(* IEC 61131-3 sources: 2026_Projet_YGO_ExcavatriceDragage/CODE_BACKUP/CODE_20260822_IntroductionTestCI/J_SUPERVISION/_BRIDGES, 7 files *)

(* ---- FB_CfgPersistBridge_BucketCfg.st ---- *)
(* =======================================================================
   💾 FB_CfgPersistBridge_BucketCfg — Pont persistance pour ST_BucketCfg
   ───────────────────────────────────────────────────────────────
   🎯 Rôle : Restauration et synchronisation bidirectionnelle IHM / Persist
   💾 Persistance : Transfert GVL_PERSISTENT <-> GVL_IHM sur Initialized
   📄 Doc métier : DOC/AF/AF_Partie-03_Contrats_Composants_v2.1.md §3
   ======================================================================= *)
FUNCTION_BLOCK FB_CfgPersistBridge_BucketCfg
VAR_OUTPUT
    // === ETATS RESTAURATION ===
    JustRestored            : BOOL;               // <-- [STAT] Vrai sur le cycle de restauration initiale
END_VAR
VAR_IN_OUT
    // === BUS CONFIGURATION ET PERSISTANCE ===
    Hmi                     : ST_BucketCfg;       // <-> [BUS] Structure de configuration IHM
    Persist                 : ST_BucketCfg;       // <-> [BUS] Structure de configuration persistante
END_VAR

JustRestored := FALSE;
IF NOT Hmi.Initialized THEN
    Hmi := Persist;
    Hmi.Initialized := TRUE;
    JustRestored := TRUE;
ELSE
    Persist := Hmi;
END_IF;

(* ---- FB_CfgPersistBridge_CommunCfg.st ---- *)
(* =======================================================================
   💾 FB_CfgPersistBridge_CommunCfg — Pont persistance pour ST_CommunCfg
   ───────────────────────────────────────────────────────────────
   🎯 Rôle : Restauration et synchronisation bidirectionnelle IHM / Persist
   💾 Persistance : Transfert GVL_PERSISTENT <-> GVL_IHM sur Initialized
   📄 Doc métier : DOC/AF/AF_Partie-03_Contrats_Composants_v2.1.md §3
   ======================================================================= *)
FUNCTION_BLOCK FB_CfgPersistBridge_CommunCfg
VAR_OUTPUT
    // === ETATS RESTAURATION ===
    JustRestored            : BOOL;               // <-- [STAT] Vrai sur le cycle de restauration initiale
END_VAR
VAR_IN_OUT
    // === BUS CONFIGURATION ET PERSISTANCE ===
    Hmi                     : ST_CommunCfg;       // <-> [BUS] Structure de configuration IHM
    Persist                 : ST_CommunCfg;       // <-> [BUS] Structure de configuration persistante
END_VAR

JustRestored := FALSE;
IF NOT Hmi.Initialized THEN
    Hmi := Persist;
    Hmi.Initialized := TRUE;
    JustRestored := TRUE;
ELSE
    Persist := Hmi;
END_IF;

(* ---- FB_CfgPersistBridge_CycleCfg.st ---- *)
(* =======================================================================
   💾 FB_CfgPersistBridge_CycleCfg — Pont persistance pour ST_CycleCfg
   ───────────────────────────────────────────────────────────────
   🎯 Rôle : Restauration et synchronisation bidirectionnelle IHM / Persist
   💾 Persistance : Transfert GVL_PERSISTENT <-> GVL_IHM sur Initialized
   📄 Doc métier : DOC/AF/AF_Partie-03_Contrats_Composants_v2.1.md §3
   ======================================================================= *)
FUNCTION_BLOCK FB_CfgPersistBridge_CycleCfg
VAR_OUTPUT
    // === ETATS RESTAURATION ===
    JustRestored            : BOOL;               // <-- [STAT] Vrai sur le cycle de restauration initiale
END_VAR
VAR_IN_OUT
    // === BUS CONFIGURATION ET PERSISTANCE ===
    Hmi                     : ST_CycleCfg;        // <-> [BUS] Structure de configuration IHM
    Persist                 : ST_CycleCfg;        // <-> [BUS] Structure de configuration persistante
END_VAR

JustRestored := FALSE;
IF NOT Hmi.Initialized THEN
    Hmi := Persist;
    Hmi.Initialized := TRUE;
    JustRestored := TRUE;
ELSE
    Persist := Hmi;
END_IF;

(* ---- FB_CfgPersistBridge_DredgingAssistCfg.st ---- *)
(* =======================================================================
   💾 FB_CfgPersistBridge_DredgingAssistCfg — Pont persistance prélèvement
   ───────────────────────────────────────────────────────────────
   🎯 Rôle : Restauration et synchronisation bidirectionnelle IHM / Persist
   💾 Persistance : Transfert GVL_PERSISTENT <-> GVL_IHM sur Initialized
   📄 Doc métier : DOC/AF/AF_Partie-03_Contrats_Composants_v2.1.md §3
   ======================================================================= *)
FUNCTION_BLOCK FB_CfgPersistBridge_DredgingAssistCfg
VAR_OUTPUT
    // === ETATS RESTAURATION ===
    JustRestored            : BOOL;               // <-- [STAT] Vrai sur le cycle de restauration initiale
END_VAR
VAR_IN_OUT
    // === BUS CONFIGURATION ET PERSISTANCE ===
    Hmi                     : ST_DredgingAssistCfg; // <-> [BUS] Structure de configuration IHM
    Persist                 : ST_DredgingAssistCfg; // <-> [BUS] Structure de configuration persistante
END_VAR

JustRestored := FALSE;
IF NOT Hmi.Initialized THEN
    Hmi := Persist;
    Hmi.Initialized := TRUE;
    JustRestored := TRUE;
ELSE
    Persist := Hmi;
END_IF;

(* ---- FB_CfgPersistBridge_SyncCfg.st ---- *)
(* =======================================================================
   💾 FB_CfgPersistBridge_SyncCfg — Pont persistance pour ST_SyncCfg
   ───────────────────────────────────────────────────────────────
   🎯 Rôle : Restauration et synchronisation bidirectionnelle IHM / Persist
   💾 Persistance : Transfert GVL_PERSISTENT <-> GVL_IHM sur Initialized
   📄 Doc métier : DOC/AF/AF_Partie-03_Contrats_Composants_v2.1.md §3
   ======================================================================= *)
FUNCTION_BLOCK FB_CfgPersistBridge_SyncCfg
VAR_OUTPUT
    // === ETATS RESTAURATION ===
    JustRestored            : BOOL;               // <-- [STAT] Vrai sur le cycle de restauration initiale
END_VAR
VAR_IN_OUT
    // === BUS CONFIGURATION ET PERSISTANCE ===
    Hmi                     : ST_SyncCfg;         // <-> [BUS] Structure de configuration IHM
    Persist                 : ST_SyncCfg;         // <-> [BUS] Structure de configuration persistante
END_VAR

JustRestored := FALSE;
IF NOT Hmi.Initialized THEN
    Hmi := Persist;
    Hmi.Initialized := TRUE;
    JustRestored := TRUE;
ELSE
    Persist := Hmi;
END_IF;

(* ---- FB_CfgPersistBridge_TranslationCfg.st ---- *)
(* =======================================================================
   💾 FB_CfgPersistBridge_TranslationCfg — Pont persistance pour ST_TranslationCfg
   ───────────────────────────────────────────────────────────────
   🎯 Rôle : Restauration et synchronisation bidirectionnelle IHM / Persist
   💾 Persistance : Transfert GVL_PERSISTENT <-> GVL_IHM sur Initialized
   📄 Doc métier : DOC/AF/AF_Partie-11_Fonction_Translation_v2.2.md
   ======================================================================= *)
FUNCTION_BLOCK FB_CfgPersistBridge_TranslationCfg
VAR_OUTPUT
    // === ETATS RESTAURATION ===
    JustRestored            : BOOL;               // <-- [STAT] Vrai sur le cycle de restauration initiale
END_VAR
VAR_IN_OUT
    // === BUS CONFIGURATION ET PERSISTANCE ===
    Hmi                     : ST_TranslationCfg;  // <-> [BUS] Structure de configuration IHM
    Persist                 : ST_TranslationCfg;  // <-> [BUS] Structure de configuration persistante
END_VAR

JustRestored := FALSE;
IF NOT Hmi.Initialized THEN
    Hmi := Persist;
    Hmi.Initialized := TRUE;
    JustRestored := TRUE;
ELSE
    Persist := Hmi;
END_IF;

(* ---- FB_CfgPersistBridge_WinchCfg.st ---- *)
(* =======================================================================
   💾 FB_CfgPersistBridge_WinchCfg — Pont persistance pour ST_WinchCfg
   ───────────────────────────────────────────────────────────────
   🎯 Rôle : Restauration et synchronisation bidirectionnelle IHM / Persist
   💾 Persistance : Transfert GVL_PERSISTENT <-> GVL_IHM sur Initialized
   📄 Doc métier : DOC/AF/AF_Partie-10_Fonction_Winch_v2.0.md
   ======================================================================= *)
FUNCTION_BLOCK FB_CfgPersistBridge_WinchCfg
VAR_OUTPUT
    // === ETATS RESTAURATION ===
    JustRestored            : BOOL;               // <-- [STAT] Vrai sur le cycle de restauration initiale
END_VAR
VAR_IN_OUT
    // === BUS CONFIGURATION ET PERSISTANCE ===
    Hmi                     : ST_WinchCfg;        // <-> [BUS] Structure de configuration IHM
    Persist                 : ST_WinchCfg;        // <-> [BUS] Structure de configuration persistante
END_VAR

JustRestored := FALSE;
IF NOT Hmi.Initialized THEN
    Hmi := Persist;
    Hmi.Initialized := TRUE;
    JustRestored := TRUE;
ELSE
    Persist := Hmi;
END_IF;
